(* PLC project PR_Gantry_2_Soft2.0 1_workflow_0f74f7_PLC, SiemensToBackhoff Siemens TIA Portal → Beckhoff TwinCAT PLCopen Converter 2.2 *)
(* stored: creationDateTime 2026-10-12T09:24:31.439330, modificationDateTime 2026-10-12T09:24:31.439330 *)

FUNCTION_BLOCK PR_Gantry_2_Soft2.0 1_workflow_0f74f7
VAR_INPUT
	iAcceptPartPick : BOOL;
	iAcceptPartPlace : BOOL;
	iAutoRunning : BOOL;
	iFaultReset : BOOL;
	iFibroSafe : BOOL;
	iOTS_Frm_Shuttle : BOOL;
	iPartPresent : BOOL;
	iPartPresent_Fibro : BOOL;
	iPartUngrip : BOOL;
	iRTR_Frm_Fibro : BOOL;
	iReset_fault : BOOL;
	iShuttleAtPickPos : BOOL;
	iShuttleSafe : BOOL;
	iSstMode : BOOL;
	iSstPB : BOOL;
	iXAxisAtPartPickPos : BOOL;
	iXAxisAtPlacePos : BOOL;
	iXAxisSafe : BOOL;
	iZAxisDownPlace : BOOL;
	iZAxisPickPos : BOOL;
	iZAxisSafe : BOOL;
	iZAxisUp : BOOL;
END_VAR
VAR_OUTPUT
	qError : ARRAY[0..8] OF BOOL;
	qMessage : ARRAY[0..1] OF BOOL;
	qOTS_To_Fibro : BOOL;
	qPartUngripCmd : BOOL;
	qRTR_To_Shuttle : BOOL;
	qXAxisHomeCmd : BOOL;
	qXAxisHomeCmdPlace : BOOL;
	qXAxisPickPosCmd : BOOL;
	qZAxisDownCmd : BOOL;
	qZAxisHomeCmd : BOOL;
	qZAxisUpCmd : BOOL;
	qZDownCmd : BOOL;
END_VAR
VAR
	c170_ChkPartPlaced_T1 : BOOL;
	c170_ChkPartPlaced_T2 : BOOL;
	c180_WtOperatorDecisionPlace_T1 : BOOL;
	c180_WtOperatorDecisionPlace_T2 : BOOL;
	c40_ChkPartPresent_T1 : BOOL;
	c40_ChkPartPresent_T2 : BOOL;
	c40_ChkPartPresent_T3 : BOOL;
	c90_ChkPartPick_T1 : BOOL;
	c90_ChkPartPick_T2 : BOOL;
	StateNo : INT;
	s100_WtOperatorDecision : BOOL;
	s100_WtOperatorDecision_T1 : BOOL;
	s100_WtOperatorDecision_T2 : BOOL;
	s10_WtAllAtSafe : BOOL;
	s10_WtAllAtSafe_T1 : BOOL;
	s110_WtZAxisUp : BOOL;
	s110_WtZAxisUp_T1 : BOOL;
	s120_ChkFibroSafe : BOOL;
	s120_ChkFibroSafe_T1 : BOOL;
	s130_WtXAxisPlacePos : BOOL;
	s130_WtXAxisPlacePos_T1 : BOOL;
	s140_WtRTRFrmFibro : BOOL;
	s140_WtRTRFrmFibro_T1 : BOOL;
	s150_WtZAxisDownPlace : BOOL;
	s150_WtZAxisDownPlace_T1 : BOOL;
	s160_WtPartUngrip : BOOL;
	s160_WtPartUngrip_T1 : BOOL;
	s170_ChkPartPlaced : BOOL;
	s170_ChkPartPlaced_T1 : BOOL;
	s170_ChkPartPlaced_T2 : BOOL;
	s180_WtOperatorDecisionPlace : BOOL;
	s180_WtOperatorDecisionPlace_T1 : BOOL;
	s180_WtOperatorDecisionPlace_T2 : BOOL;
	s1_ResetRelease : BOOL;
	s1_ResetRelease_T1 : BOOL;
	s20_WtZAxisSafe : BOOL;
	s20_WtZAxisSafe_T1 : BOOL;
	s30_WtXAxisAtSafe : BOOL;
	s30_WtXAxisAtSafe_T1 : BOOL;
	s40_ChkPartPresent : BOOL;
	s40_ChkPartPresent_T1 : BOOL;
	s40_ChkPartPresent_T2 : BOOL;
	s40_ChkPartPresent_T3 : BOOL;
	s45_WtOperatorAck : BOOL;
	s45_WtOperatorAck_T1 : BOOL;
	s50_WtShuttleAtSafe : BOOL;
	s50_WtShuttleAtSafe_T1 : BOOL;
	s60_WtXAxisPickPos : BOOL;
	s60_WtXAxisPickPos_T1 : BOOL;
	s70_WtOTSFrmShuttle : BOOL;
	s70_WtOTSFrmShuttle_T1 : BOOL;
	s80_WtZAxisPickPos : BOOL;
	s80_WtZAxisPickPos_T1 : BOOL;
	s90_ChkPartPick : BOOL;
	s90_ChkPartPick_T1 : BOOL;
	s90_ChkPartPick_T2 : BOOL;
	sAbnormalStatus : BOOL;
	sPartPresentInGrip : BOOL;
	sSst : BOOL;
	sSstPulse : BOOL;
	sSstRise : R_TRIG;
	sStWtResetRel : BOOL;
	sStWtResetRel_T1 : BOOL;
END_VAR
VAR_TEMP
	tOne : BOOL;
END_VAR
  VAR  (* added by the conversion: wires and edge detectors of the diagram *)
    _w24 : BOOL;
    _w26 : BOOL;
    _w39 : BOOL;
    _w41 : BOOL;
    _w42 : BOOL;
    _w56 : BOOL;
    _w58 : BOOL;
    _w59 : BOOL;
    _w72 : BOOL;
    _w74 : BOOL;
    _w75 : BOOL;
    _w92 : BOOL;
    _w96 : BOOL;
    _w97 : BOOL;
    _w133 : BOOL;
    _w136 : BOOL;
    _w137 : BOOL;
    _w138 : BOOL;
    _w139 : BOOL;
    _w152 : BOOL;
    _w154 : BOOL;
    _w155 : BOOL;
    _w172 : BOOL;
    _w174 : BOOL;
    _w175 : BOOL;
    _w188 : BOOL;
    _w190 : BOOL;
    _w191 : BOOL;
    _w208 : BOOL;
    _w210 : BOOL;
    _w211 : BOOL;
    _w228 : BOOL;
    _w230 : BOOL;
    _w231 : BOOL;
    _w269 : BOOL;
    _w272 : BOOL;
    _w273 : BOOL;
    _w274 : BOOL;
    _w294 : BOOL;
    _w296 : BOOL;
    _w297 : BOOL;
    _w298 : BOOL;
    _w316 : BOOL;
    _w320 : BOOL;
    _w321 : BOOL;
    _w338 : BOOL;
    _w340 : BOOL;
    _w341 : BOOL;
    _w354 : BOOL;
    _w356 : BOOL;
    _w357 : BOOL;
    _w374 : BOOL;
    _w376 : BOOL;
    _w377 : BOOL;
    _w394 : BOOL;
    _w396 : BOOL;
    _w397 : BOOL;
    _w414 : BOOL;
    _w416 : BOOL;
    _w417 : BOOL;
    _w449 : BOOL;
    _w452 : BOOL;
    _w453 : BOOL;
    _w454 : BOOL;
    _w482 : BOOL;
    _w484 : BOOL;
    _w485 : BOOL;
    _w486 : BOOL;
  END_VAR

(* LD diagram, written out as Structured Text *)
(* Network 1 *)
(* Create Single Step Pulse bit *)
(* Create Single Step bit *)
(* Transition for STATE Num:0 Reset Released *)
(* STATE Num:0 Reset Released *)
(* Transition for STATE Num:1 ResetRelease *)
(* STATE Num:1 ResetRelease *)
(* Transition for STATE Num:10 WtAllAtSafe *)
(* STATE Num:10 WtAllAtSafe *)
(* Transition for STATE Num:20 WtZAxisSafe *)
(* STATE Num:20 WtZAxisSafe *)
(* Actions for STATE Num:20 WtZAxisSafe *)
(* Transition for STATE Num:30 WtXAxisAtSafe *)
(* STATE Num:30 WtXAxisAtSafe *)
(* Actions for STATE Num:30 WtXAxisAtSafe *)
(* Condition1 for STATE Num:40 ChkPartPresent *)
(* Condition2 for STATE Num:40 ChkPartPresent *)
(* Condition3 for STATE Num:40 ChkPartPresent *)
(* Transition for STATE Num:40 ChkPartPresent *)
(* STATE Num:40 ChkPartPresent *)
(* Transition for STATE Num:45 WtOperatorAck *)
(* STATE Num:45 WtOperatorAck *)
(* Actions for STATE Num:45 WtOperatorAck *)
(* Transition for STATE Num:50 WtShuttleAtSafe *)
(* STATE Num:50 WtShuttleAtSafe *)
(* Transition for STATE Num:60 WtXAxisPickPos *)
(* STATE Num:60 WtXAxisPickPos *)
(* Actions for STATE Num:60 WtXAxisPickPos *)
(* Transition for STATE Num:70 WtOTSFrmShuttle *)
(* STATE Num:70 WtOTSFrmShuttle *)
(* Actions for STATE Num:70 WtOTSFrmShuttle *)
(* Transition for STATE Num:80 WtZAxisPickPos *)
(* STATE Num:80 WtZAxisPickPos *)
(* Actions for STATE Num:80 WtZAxisPickPos - qZAxisDownCmd *)
(* Actions for STATE Num:80 WtZAxisPickPos - qError[5] on condition *)
(* Condition1 for STATE Num:90 ChkPartPick *)
(* Condition2 for STATE Num:90 ChkPartPick *)
(* Transition for STATE Num:90 ChkPartPick *)
(* STATE Num:90 ChkPartPick *)
(* Actions for STATE Num:90 ChkPartPick - qError[3] on Condition1 *)
(* Transition for STATE Num:100 WtOperatorDecision *)
(* STATE Num:100 WtOperatorDecision *)
(* Actions for STATE Num:100 WtOperatorDecision *)
(* Transition for STATE Num:110 WtZAxisUp *)
(* STATE Num:110 WtZAxisUp *)
(* Actions for STATE Num:110 WtZAxisUp *)
(* Transition for STATE Num:120 ChkFibroSafe *)
(* STATE Num:120 ChkFibroSafe *)
(* Transition for STATE Num:130 WtXAxisPlacePos *)
(* STATE Num:130 WtXAxisPlacePos *)
(* Actions for STATE Num:130 WtXAxisPlacePos *)
(* Transition for STATE Num:140 WtRTRFrmFibro *)
(* STATE Num:140 WtRTRFrmFibro *)
(* Actions for STATE Num:140 WtRTRFrmFibro *)
(* Transition for STATE Num:150 WtZAxisDownPlace *)
(* STATE Num:150 WtZAxisDownPlace *)
(* Actions for STATE Num:150 WtZAxisDownPlace *)
(* Transition for STATE Num:160 WtPartUngrip *)
(* STATE Num:160 WtPartUngrip *)
(* Actions for STATE Num:160 WtPartUngrip *)
(* Condition1 for STATE Num:170 ChkPartPlaced *)
(* Condition2 for STATE Num:170 ChkPartPlaced *)
(* Transition for STATE Num:170 ChkPartPlaced *)
(* STATE Num:170 ChkPartPlaced *)
(* Actions for STATE Num:170 ChkPartPlaced *)
(* Condition1 for STATE Num:180 WtOperatorDecisionPlace *)
(* Condition2 for STATE Num:180 WtOperatorDecisionPlace *)
(* Transition for STATE Num:180 WtOperatorDecisionPlace *)
(* STATE Num:180 WtOperatorDecisionPlace *)
(* Actions for STATE Num:180 WtOperatorDecisionPlace *)
tOne := tOne OR NOT tOne;
sSstRise(CLK := iSstPB);
sSstPulse := sSstRise.Q;
sSst := iSstMode AND sSstPulse OR NOT iSstMode;
sStWtResetRel_T1 := sStWtResetRel AND iAutoRunning;
_w24 := sStWtResetRel;
_w26 := (_w24 OR NOT iAutoRunning) AND NOT sStWtResetRel_T1;
sStWtResetRel := _w26;
IF _w26 THEN StateNo := 0; END_IF;
s1_ResetRelease_T1 := s1_ResetRelease AND NOT sStWtResetRel AND sSst AND iAutoRunning;
_w39 := s1_ResetRelease;
_w41 := (_w39 OR sStWtResetRel_T1) AND NOT sStWtResetRel;
_w42 := _w41 AND NOT s1_ResetRelease_T1;
s1_ResetRelease := _w42;
IF _w42 THEN StateNo := 1; END_IF;
s10_WtAllAtSafe_T1 := s10_WtAllAtSafe AND NOT sStWtResetRel AND sSst AND iShuttleSafe AND iFibroSafe;
_w56 := s10_WtAllAtSafe;
_w58 := (_w56 OR s1_ResetRelease_T1) AND NOT sStWtResetRel;
_w59 := _w58 AND NOT s10_WtAllAtSafe_T1;
s10_WtAllAtSafe := _w59;
IF _w59 THEN StateNo := 10; END_IF;
s20_WtZAxisSafe_T1 := s20_WtZAxisSafe AND NOT sStWtResetRel AND sSst AND iZAxisSafe;
_w72 := s20_WtZAxisSafe;
_w74 := (_w72 OR s10_WtAllAtSafe_T1) AND NOT sStWtResetRel;
_w75 := _w74 AND NOT s20_WtZAxisSafe_T1;
s20_WtZAxisSafe := _w75;
IF _w75 THEN StateNo := 20; END_IF;
qZAxisHomeCmd := s20_WtZAxisSafe;
s30_WtXAxisAtSafe_T1 := s30_WtXAxisAtSafe AND NOT sStWtResetRel AND sSst AND iXAxisSafe;
_w92 := s30_WtXAxisAtSafe;
_w96 := (_w92 OR s180_WtOperatorDecisionPlace_T1 OR s170_ChkPartPlaced_T2 OR s20_WtZAxisSafe_T1) AND NOT sStWtResetRel;
_w97 := _w96 AND NOT s30_WtXAxisAtSafe_T1;
s30_WtXAxisAtSafe := _w97;
IF _w97 THEN StateNo := 30; END_IF;
qXAxisHomeCmd := s30_WtXAxisAtSafe;
c40_ChkPartPresent_T1 := sAbnormalStatus;
c40_ChkPartPresent_T2 := iPartPresent;
c40_ChkPartPresent_T3 := NOT iPartPresent;
s40_ChkPartPresent_T1 := s40_ChkPartPresent AND NOT sStWtResetRel AND sSst AND c40_ChkPartPresent_T1;
s40_ChkPartPresent_T2 := s40_ChkPartPresent AND NOT sStWtResetRel AND sSst AND NOT s40_ChkPartPresent_T1 AND c40_ChkPartPresent_T2;
s40_ChkPartPresent_T3 := s40_ChkPartPresent AND NOT sStWtResetRel AND sSst AND NOT s40_ChkPartPresent_T1 AND NOT s40_ChkPartPresent_T1 AND NOT s40_ChkPartPresent_T2 AND c40_ChkPartPresent_T3;
_w133 := s40_ChkPartPresent;
_w136 := (_w133 OR s45_WtOperatorAck_T1 OR s30_WtXAxisAtSafe_T1) AND NOT sStWtResetRel;
_w137 := _w136 AND NOT s40_ChkPartPresent_T1;
_w138 := _w137 AND NOT s40_ChkPartPresent_T2;
_w139 := _w138 AND NOT s40_ChkPartPresent_T3;
s40_ChkPartPresent := _w139;
IF _w139 THEN StateNo := 40; END_IF;
s45_WtOperatorAck_T1 := s45_WtOperatorAck AND NOT sStWtResetRel AND sSst AND iFaultReset;
_w152 := s45_WtOperatorAck;
_w154 := (_w152 OR s40_ChkPartPresent_T1) AND NOT sStWtResetRel;
_w155 := _w154 AND NOT s45_WtOperatorAck_T1;
s45_WtOperatorAck := _w155;
IF _w155 THEN StateNo := 45; END_IF;
qError[8] := s45_WtOperatorAck;
s50_WtShuttleAtSafe_T1 := s50_WtShuttleAtSafe AND NOT sStWtResetRel AND sSst AND iShuttleSafe;
_w172 := s50_WtShuttleAtSafe;
_w174 := (_w172 OR s40_ChkPartPresent_T3) AND NOT sStWtResetRel;
_w175 := _w174 AND NOT s50_WtShuttleAtSafe_T1;
s50_WtShuttleAtSafe := _w175;
IF _w175 THEN StateNo := 50; END_IF;
s60_WtXAxisPickPos_T1 := s60_WtXAxisPickPos AND NOT sStWtResetRel AND sSst AND iXAxisAtPartPickPos;
_w188 := s60_WtXAxisPickPos;
_w190 := (_w188 OR s50_WtShuttleAtSafe_T1) AND NOT sStWtResetRel;
_w191 := _w190 AND NOT s60_WtXAxisPickPos_T1;
s60_WtXAxisPickPos := _w191;
IF _w191 THEN StateNo := 60; END_IF;
qXAxisPickPosCmd := s60_WtXAxisPickPos;
s70_WtOTSFrmShuttle_T1 := s70_WtOTSFrmShuttle AND NOT sStWtResetRel AND sSst AND iOTS_Frm_Shuttle;
_w208 := s70_WtOTSFrmShuttle;
_w210 := (_w208 OR s60_WtXAxisPickPos_T1) AND NOT sStWtResetRel;
_w211 := _w210 AND NOT s70_WtOTSFrmShuttle_T1;
s70_WtOTSFrmShuttle := _w211;
IF _w211 THEN StateNo := 70; END_IF;
qRTR_To_Shuttle := s70_WtOTSFrmShuttle;
s80_WtZAxisPickPos_T1 := s80_WtZAxisPickPos AND NOT sStWtResetRel AND sSst AND iZAxisPickPos;
_w228 := s80_WtZAxisPickPos;
_w230 := (_w228 OR s70_WtOTSFrmShuttle_T1) AND NOT sStWtResetRel;
_w231 := _w230 AND NOT s80_WtZAxisPickPos_T1;
s80_WtZAxisPickPos := _w231;
IF _w231 THEN StateNo := 80; END_IF;
qZAxisDownCmd := s80_WtZAxisPickPos;
qError[5] := s80_WtZAxisPickPos AND qZAxisDownCmd AND NOT iShuttleAtPickPos;
c90_ChkPartPick_T1 := iPartPresent AND NOT sPartPresentInGrip OR NOT iPartPresent AND sPartPresentInGrip;
c90_ChkPartPick_T2 := NOT iPartPresent AND sPartPresentInGrip;
s90_ChkPartPick_T1 := s90_ChkPartPick AND NOT sStWtResetRel AND sSst AND c90_ChkPartPick_T1;
s90_ChkPartPick_T2 := s90_ChkPartPick AND NOT sStWtResetRel AND sSst AND NOT s90_ChkPartPick_T1 AND c90_ChkPartPick_T2;
_w269 := s90_ChkPartPick;
_w272 := (_w269 OR s100_WtOperatorDecision_T2 OR s80_WtZAxisPickPos_T1) AND NOT sStWtResetRel;
_w273 := _w272 AND NOT s90_ChkPartPick_T1;
_w274 := _w273 AND NOT s90_ChkPartPick_T2;
s90_ChkPartPick := _w274;
IF _w274 THEN StateNo := 90; END_IF;
qError[3] := s90_ChkPartPick_T1;
s100_WtOperatorDecision_T1 := s100_WtOperatorDecision AND NOT sStWtResetRel AND sSst AND iAcceptPartPick;
s100_WtOperatorDecision_T2 := s100_WtOperatorDecision AND NOT sStWtResetRel AND sSst AND NOT s100_WtOperatorDecision_T1 AND iFaultReset;
_w294 := s100_WtOperatorDecision;
_w296 := (_w294 OR s90_ChkPartPick_T1) AND NOT sStWtResetRel;
_w297 := _w296 AND NOT s100_WtOperatorDecision_T1;
_w298 := _w297 AND NOT s100_WtOperatorDecision_T2;
s100_WtOperatorDecision := _w298;
IF _w298 THEN StateNo := 100; END_IF;
qError[1] := s100_WtOperatorDecision;
qMessage[0] := s100_WtOperatorDecision;
s110_WtZAxisUp_T1 := s110_WtZAxisUp AND NOT sStWtResetRel AND sSst AND iZAxisUp;
_w316 := s110_WtZAxisUp;
_w320 := (_w316 OR s100_WtOperatorDecision_T1 OR s90_ChkPartPick_T2 OR s40_ChkPartPresent_T2) AND NOT sStWtResetRel;
_w321 := _w320 AND NOT s110_WtZAxisUp_T1;
s110_WtZAxisUp := _w321;
IF _w321 THEN StateNo := 110; END_IF;
qZAxisUpCmd := s110_WtZAxisUp;
s120_ChkFibroSafe_T1 := s120_ChkFibroSafe AND NOT sStWtResetRel AND sSst AND iFibroSafe;
_w338 := s120_ChkFibroSafe;
_w340 := (_w338 OR s110_WtZAxisUp_T1) AND NOT sStWtResetRel;
_w341 := _w340 AND NOT s120_ChkFibroSafe_T1;
s120_ChkFibroSafe := _w341;
IF _w341 THEN StateNo := 120; END_IF;
s130_WtXAxisPlacePos_T1 := s130_WtXAxisPlacePos AND NOT sStWtResetRel AND sSst AND iXAxisAtPlacePos;
_w354 := s130_WtXAxisPlacePos;
_w356 := (_w354 OR s120_ChkFibroSafe_T1) AND NOT sStWtResetRel;
_w357 := _w356 AND NOT s130_WtXAxisPlacePos_T1;
s130_WtXAxisPlacePos := _w357;
IF _w357 THEN StateNo := 130; END_IF;
qXAxisHomeCmdPlace := s130_WtXAxisPlacePos;
s140_WtRTRFrmFibro_T1 := s140_WtRTRFrmFibro AND NOT sStWtResetRel AND sSst AND iRTR_Frm_Fibro;
_w374 := s140_WtRTRFrmFibro;
_w376 := (_w374 OR s130_WtXAxisPlacePos_T1) AND NOT sStWtResetRel;
_w377 := _w376 AND NOT s140_WtRTRFrmFibro_T1;
s140_WtRTRFrmFibro := _w377;
IF _w377 THEN StateNo := 140; END_IF;
qOTS_To_Fibro := s140_WtRTRFrmFibro;
s150_WtZAxisDownPlace_T1 := s150_WtZAxisDownPlace AND NOT sStWtResetRel AND sSst AND iZAxisDownPlace;
_w394 := s150_WtZAxisDownPlace;
_w396 := (_w394 OR s140_WtRTRFrmFibro_T1) AND NOT sStWtResetRel;
_w397 := _w396 AND NOT s150_WtZAxisDownPlace_T1;
s150_WtZAxisDownPlace := _w397;
IF _w397 THEN StateNo := 150; END_IF;
qZDownCmd := s150_WtZAxisDownPlace;
s160_WtPartUngrip_T1 := s160_WtPartUngrip AND NOT sStWtResetRel AND sSst AND iPartUngrip;
_w414 := s160_WtPartUngrip;
_w416 := (_w414 OR s150_WtZAxisDownPlace_T1) AND NOT sStWtResetRel;
_w417 := _w416 AND NOT s160_WtPartUngrip_T1;
s160_WtPartUngrip := _w417;
IF _w417 THEN StateNo := 160; END_IF;
qPartUngripCmd := s160_WtPartUngrip;
c170_ChkPartPlaced_T1 := iPartPresent AND NOT sPartPresentInGrip OR NOT iPartPresent AND sPartPresentInGrip;
c170_ChkPartPlaced_T2 := iPartPresent_Fibro AND NOT sPartPresentInGrip;
s170_ChkPartPlaced_T1 := s170_ChkPartPlaced AND NOT sStWtResetRel AND sSst AND c170_ChkPartPlaced_T1;
s170_ChkPartPlaced_T2 := s170_ChkPartPlaced AND NOT sStWtResetRel AND sSst AND NOT s170_ChkPartPlaced_T1 AND c170_ChkPartPlaced_T2;
_w449 := s170_ChkPartPlaced;
_w452 := (_w449 OR s180_WtOperatorDecisionPlace_T2 OR s160_WtPartUngrip_T1) AND NOT sStWtResetRel;
_w453 := _w452 AND NOT s170_ChkPartPlaced_T1;
_w454 := _w453 AND NOT s170_ChkPartPlaced_T2;
s170_ChkPartPlaced := _w454;
IF _w454 THEN StateNo := 170; END_IF;
qError[3] := s170_ChkPartPlaced;
c180_WtOperatorDecisionPlace_T1 := iAcceptPartPlace;
c180_WtOperatorDecisionPlace_T2 := iFaultReset;
s180_WtOperatorDecisionPlace_T1 := s180_WtOperatorDecisionPlace AND NOT sStWtResetRel AND sSst AND c180_WtOperatorDecisionPlace_T1;
s180_WtOperatorDecisionPlace_T2 := s180_WtOperatorDecisionPlace AND NOT sStWtResetRel AND sSst AND NOT s180_WtOperatorDecisionPlace_T1 AND c180_WtOperatorDecisionPlace_T2;
_w482 := s180_WtOperatorDecisionPlace;
_w484 := (_w482 OR s170_ChkPartPlaced_T1) AND NOT sStWtResetRel;
_w485 := _w484 AND NOT s180_WtOperatorDecisionPlace_T1;
_w486 := _w485 AND NOT s180_WtOperatorDecisionPlace_T2;
s180_WtOperatorDecisionPlace := _w486;
IF _w486 THEN StateNo := 180; END_IF;
qMessage[1] := s180_WtOperatorDecisionPlace;
qError[2] := s180_WtOperatorDecisionPlace;
END_FUNCTION_BLOCK
